// Mitsubishi GX Works2 project: 시험1_단속동작   PLC: FX3U/FX3UC

PROGRAM MAIN
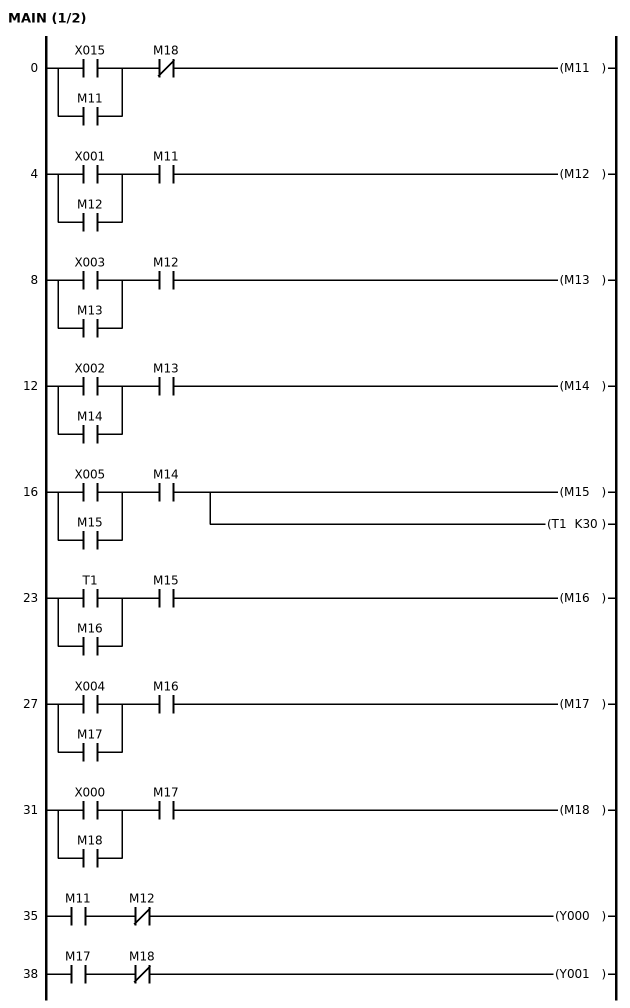
0     LD      X015
      OR      M11
      ANI     M18
      OUT     M11
4     LD      X001
      OR      M12
      AND     M11
      OUT     M12
8     LD      X003
      OR      M13
      AND     M12
      OUT     M13
12    LD      X002
      OR      M14
      AND     M13
      OUT     M14
16    LD      X005
      OR      M15
      AND     M14
      OUT     M15
      OUT     T1 K30
23    LD      T1
      OR      M16
      AND     M15
      OUT     M16
27    LD      X004
      OR      M17
      AND     M16
      OUT     M17
31    LD      X000
      OR      M18
      AND     M17
      OUT     M18
35    LD      M11
      ANI     M12
      OUT     Y000
38    LD      M17
      ANI     M18
      OUT     Y001
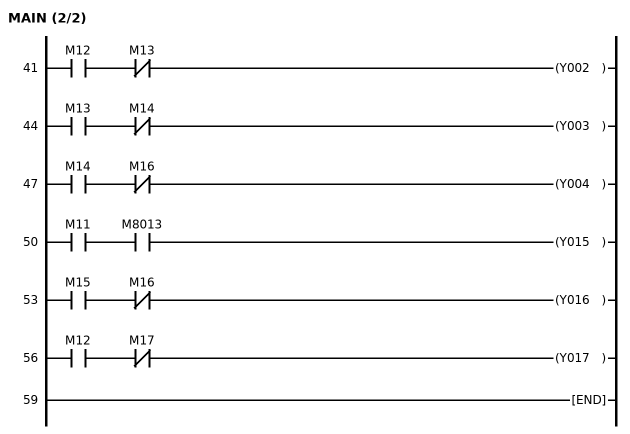
41    LD      M12
      ANI     M13
      OUT     Y002
44    LD      M13
      ANI     M14
      OUT     Y003
47    LD      M14
      ANI     M16
      OUT     Y004
50    LD      M11
      AND     M8013
      OUT     Y015
53    LD      M15
      ANI     M16
      OUT     Y016
56    LD      M12
      ANI     M17
      OUT     Y017
59    END
END_PROGRAM
